// TwinCAT 3 PLC project PLCStudent
// ProgramVersion: 3.1.4026.20
// libraries:
//   Tc2_Standard, * (Beckhoff Automation GmbH)
//   Tc2_System, * (Beckhoff Automation GmbH)
//   Tc3_Module, * (Beckhoff Automation GmbH)
// project tree:
//   / PlcTask.TcTTO
//   POUs/ MAIN.TcPOU, Control_FBD.TcPOU
// (motion and I/O tree: see PLC project plcsim)
// real-time tasks:
//   TASK PlcTask: cycle T#80ms, priority 1, ADS port 350
//   TASK PlcTask1: cycle T#10ms, priority 20, ADS port 351
// variable links:
//   PLCSim/PLCSim Instance <-> PLCStudent/PLCStudent Instance
//     PlcTask Inputs/GVL.ixBack <-> PlcTask Outputs/Control_FBD.qxBack
//     PlcTask Inputs/GVL.ixDispBit1 <-> PlcTask Outputs/Control_FBD.qxDispBit1
//     PlcTask Inputs/GVL.ixDispBit2 <-> PlcTask Outputs/Control_FBD.qxDispBit2
//     PlcTask Inputs/GVL.ixDrain <-> PlcTask Outputs/Control_FBD.qxDrain
//     PlcTask Inputs/GVL.ixFill <-> PlcTask Outputs/Control_FBD.qxFill
//     PlcTask Inputs/GVL.ixForw <-> PlcTask Outputs/Control_FBD.qxForw
//     PlcTask Inputs/GVL.ixHeat <-> PlcTask Outputs/Control_FBD.qxHeat
//     PlcTask Inputs/GVL.ixSpin <-> PlcTask Outputs/Control_FBD.qxSpin
//     PlcTask Outputs/GVL.qxLevel1 <-> PlcTask Inputs/Control_FBD.ixLevel1
//     PlcTask Outputs/GVL.qxLevel2 <-> PlcTask Inputs/Control_FBD.ixLevel2
//     PlcTask Outputs/GVL.qxLevel3 <-> PlcTask Inputs/Control_FBD.ixLevel3
//     PlcTask Outputs/GVL.qxNotEmpty <-> PlcTask Inputs/Control_FBD.ixNotEmpty
//     PlcTask Outputs/GVL.qxPulse <-> PlcTask Inputs/Control_FBD.ixPulse
//     PlcTask Outputs/GVL.qxSetLevel <-> PlcTask Inputs/Control_FBD.ixSetLevel
//     PlcTask Outputs/GVL.qxStart <-> PlcTask Inputs/Control_FBD.ixStart
//     PlcTask Outputs/GVL.qxTempOk <-> PlcTask Inputs/Control_FBD.ixTempOk

CONFIGURATION PLCStudent
    RESOURCE PLC ON TwinCAT3
        TASK PlcTask(INTERVAL := T#10ms, PRIORITY := 20);
        PROGRAM MAIN WITH PlcTask : MAIN;
    END_RESOURCE
END_CONFIGURATION

// ---- POUs/MAIN.TcPOU
PROGRAM MAIN
VAR
END_VAR

Control_FBD();

END_PROGRAM

// ---- POUs/Control_FBD.TcPOU
PROGRAM Control_FBD
VAR
	
	ixPulse			AT %I*:	BOOL; 		(* PULS button *)
	ixStart			AT %I*:	BOOL; 		(* START switch *)
	ixSetLevel		AT %I*:	BOOL; 		(* NIVÅ switch *)
	ixLevel3		AT %I*:	BOOL; 		(* Sensor for level 3 *)
	ixLevel2		AT %I*:	BOOL; 		(* Sensor for level 2 *)
	ixLevel1		AT %I*:	BOOL; 		(* Sensor for level 1 *)
	ixNotEmpty		AT %I*:	BOOL; 		(* Sensor for not empty *)
	ixTempOk		AT %I*:	BOOL; 		(* Temp sensor *)
	
	mxFill : BOOL;
	mxForw : BOOL;
	mxBack : BOOL;
	mxSpin : BOOL;
	mxDrain : BOOL;
	mxHeat : BOOL;
	
	qxForw			AT %Q*:	BOOL; 		(* Washer cylinder forward *)
	qxBack			AT %Q*:	BOOL; 		(* Washer cylinder back *)
	qxSpin			AT %Q*:	BOOL; 		(* Hi-spin/Centrifuge need qxForw or qxBack*)
	qxFill			AT %Q*:	BOOL; 		(* Fill water *)
	qxDrain			AT %Q*:	BOOL; 		(* Drain water *)
	qxHeat			AT %Q*:	BOOL; 		(* Heat water *)
	qxDispBit1		AT %Q*:	BOOL; 		(* Display bit 1 *)
	qxDispBit2		AT %Q*:	BOOL; 		(* Display bit 2 *)
END_VAR

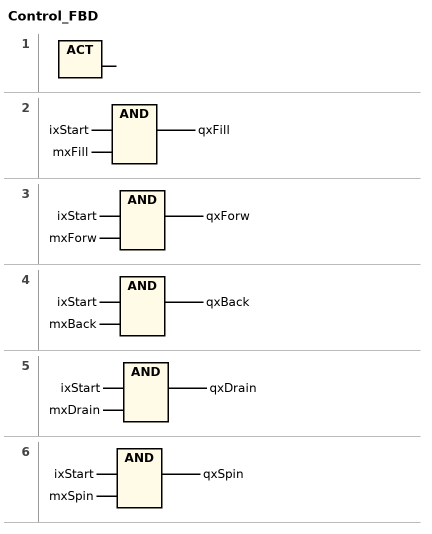
// NETWORK 1
ACT();

// NETWORK 2
qxFill := ixStart AND mxFill;

// NETWORK 3
qxForw := ixStart AND mxForw;

// NETWORK 4
qxBack := ixStart AND mxBack;

// NETWORK 5
qxDrain := ixStart AND mxDrain;

// NETWORK 6
qxSpin := ixStart AND mxSpin;

ACTION ACT:
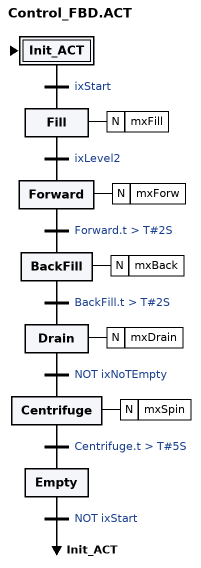
INITIAL_STEP Init_ACT:
END_STEP
TRANSITION FROM Init_ACT TO Fill
    := ixStart;
END_TRANSITION
STEP Fill:
    mxFill(N);
END_STEP
TRANSITION FROM Fill TO Forward
    := ixLevel2;
END_TRANSITION
STEP Forward:
    mxForw(N);
END_STEP
TRANSITION FROM Forward TO BackFill
    := Forward.t > T#2S;
END_TRANSITION
STEP BackFill:
    mxBack(N);
END_STEP
TRANSITION FROM BackFill TO Drain
    := BackFill.t > T#2S;
END_TRANSITION
STEP Drain:
    mxDrain(N);
END_STEP
TRANSITION FROM Drain TO Centrifuge
    := NOT ixNoTEmpty;
END_TRANSITION
STEP Centrifuge:
    mxSpin(N);
END_STEP
TRANSITION FROM Centrifuge TO Empty
    := Centrifuge.t > T#5S;
END_TRANSITION
STEP Empty:
END_STEP
TRANSITION FROM Empty TO Init_ACT
    := NOT ixStart;
END_TRANSITION
END_ACTION

END_PROGRAM
